// TIA Portal V21 export
FUNCTION "Enable" : Bool   // FC2, F_LAD
{ S7_Optimized_Access := 'TRUE' }
// True while both inputs are true.
   VAR_INPUT
      "a" : Bool;
      "b" : Bool;
   END_VAR
BEGIN

REGION Network 1: Both inputs
   // On while both inputs are on.
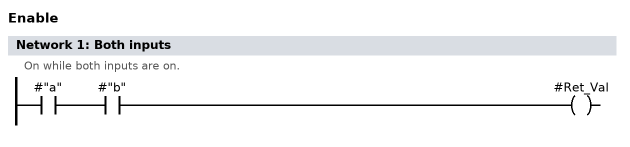
   RUNG wire#powerrail
      Contact( #"a" )
      Contact( #"b" )
      Coil( #Ret_Val )
   END_RUNG
   // the same network as SCL:
   #Ret_Val := #"a" AND #"b";
END_REGION
END_FUNCTION
